Staubli VAL3: tx2.pjx

--- tx2.pjx ---
Parameters version=s8.10.5Cs9_BS2172 stackSize=20000 millimeterUnit=true
Program file=getPath.pgx
Program file=initArmInfo.pgx
Program file=initDataBase.pgx
Program file=initWidget.pgx
Program file=mainCycle.pgx
Program file=moveCalPos.pgx
Program file=moveRecPos.pgx
Program file=refreshBtn0_CaliTcp.pgx
Program file=refreshBtn1_AdjXY.pgx
Program file=refreshBtn2_AdjZ.pgx
Program file=refreshBtn3_Test.pgx
Program file=saveCall.pgx
Program file=saveTask.pgx
Program file=start.pgx
Program file=stop.pgx
Data file=tx2.dtx
Library alias=algorithm path=Disk://SmartTCP_CS9/Algorithm6/Algorithm6.pjx
Library alias=db path=Disk://SmartTCP_CS9/DataBase6/DataBase6.pjx

--- tx2.dtx ---


--- start.pgx ---
public program start()
begin
  call initArmInfo()
  call initWidget()
  call initDataBase()
  call mainCycle()
end

--- getPath.pgx ---
program getPath(string x_sHmiName, string& x_sHmiPath)
begin
  x_sHmiPath=libPath()+"/interface/"+x_sHmiName
end

--- initArmInfo.pgx ---
program initArmInfo()
  local string l_sLanguage
  local string l_sMounting
begin
  //*******************************************************
  db:utLbl_Axis_Data.Common.sText="6axis"
  //*******************************************************
  //Get mounting property
  //*******************************************************
  l_sMounting=getVersion("Arm Mounting")
  switch l_sMounting
    case "floor"
      db:sMounting="Floor"
      db:utCbx_Mounting_Data.Common.sValue="Floor"
    break
    case "ceiling"
      db:sMounting="Ceiling"
      db:utCbx_Mounting_Data.Common.sValue="Ceiling"
    break
    default
      db:sMounting="Null"
      db:utCbx_Mounting_Data.Common.sValue=""
    break
  endSwitch
  //*******************************************************
  //Get system language
  //*******************************************************
  l_sLanguage=getLanguage()
  switch l_sLanguage
    case "chinese"
      db:sLanguage="chinese"
      db:utCbx_Language_Data.Common.sValue="Chinese"
    break
    case "english"
      db:sLanguage="english"
      db:utCbx_Language_Data.Common.sValue="English"
    break
    default
      db:sLanguage="english"
      db:utCbx_Language_Data.Common.sValue="English"
    break
  endSwitch
  //
  //*******************************************************
  //Initialize the flange as the current tool
  //*******************************************************
  call db:updateTool(0,false)
end

--- initDataBase.pgx ---
program initDataBase()
begin
  db:nStep0=10
  db:nStep1=10
  db:nStep2=10
  db:nStep3=10
  //
  db:tFlange.trsf={0,0,0,0,0,0}
  db:trOffset={0,0,10,0,0,0}
  //
  db:mSpeed_C_blend.tvel=250
  db:mSpeed_C_blend.blend=Cartesian
  db:mSpeed_C_blend.leave=0
  db:mSpeed_C_blend.reach=0
  //
  db:mSpeed_J_blend.tvel=250
  db:mSpeed_J_blend.blend=joint
  db:mSpeed_J_blend.leave=5
  db:mSpeed_J_blend.reach=5
  //
  db:mSlow.tvel=30
  db:mSlow.blend=Cartesian
  db:mSlow.leave=0
  db:mSlow.reach=0
  //
  db:cConfigSame={ssame,esame,wsame}
  //
  //pTeach1.trsf={0,0,0,0,0,0}
  db:pTeach1.config={ssame,esame,wsame}
  //pTeach2.trsf={0,0,0,0,0,0}
  db:pTeach2.config={ssame,esame,wsame}
  //pTeach3.trsf={0,0,0,0,0,0}
  db:pTeach3.config={ssame,esame,wsame}
  //pTeach4.trsf={0,0,0,0,0,0}
  db:pTeach4.config={ssame,esame,wsame}
  //pTeach5.trsf={0,0,0,0,0,0}
  db:pTeach5.config={ssame,esame,wsame}
  //pTeach6.trsf={0,0,0,0,0,0}
  db:pTeach6.config={ssame,esame,wsame}
  //pTeach6.trsf={0,0,0,0,0,0}
  db:pTeach7.config={ssame,esame,wsame}
  //
  //pAdjustXY_2_1.trsf={0,0,0,0,0,0}
  db:pAdjustXY_2_1.config={ssame,esame,wsame}
  //pAdjustXY_2_2.trsf={0,0,0,0,0,0}
  db:pAdjustXY_2_2.config={ssame,esame,wsame}
  //pAdjustXY_3_1.trsf={0,0,0,0,0,0}
  db:pAdjustXY_3_1.config={ssame,esame,wsame}
  //pAdjustXY_3_2.trsf={0,0,0,0,0,0}
  db:pAdjustXY_3_2.config={ssame,esame,wsame}
  //pAdjustXY_3_3.trsf={0,0,0,0,0,0}
  db:pAdjustXY_3_3.config={ssame,esame,wsame}
  //pAdjustZ_2_1.trsf={0,0,0,0,0,0}
  db:pAdjustZ_2_1.config={ssame,esame,wsame}
  //pAdjustZ_2_2.trsf={0,0,0,0,0,0}
  db:pAdjustZ_2_2.config={ssame,esame,wsame}
  //
  db:bTeach1=false
  db:bTeach2=false
  db:bTeach3=false
  db:bTeach4=false
  db:bTeach5=false
  db:bTeach6=false
  db:bTeach7=false
  //
  db:bAdjustXY_2_1=false
  db:bAdjustXY_2_2=false
  db:bAdjustXY_3_1=false
  db:bAdjustXY_3_2=false
  db:bAdjustXY_3_3=false
  db:bAdjustZ_2_1=false
  db:bAdjustZ_2_2=false
  //
  db:sLanguageM=""
  db:sCbxLanguage=""
  db:sCbxMounting=""
end

--- initWidget.pgx ---
program initWidget()
  local num l_nI
  local string l_sID
  local string l_sPage
begin
  //*************************************************************************************************
  //Initialize the widgets of the <Page_Main>：
  //*************************************************************************************************
  call getPath("Page_Main",l_sPage)
  //Container
  call db:initContainer(db:utCtn_Function,l_sPage,"ctn_Function",true)
  db:utCtn_Function.Common.sSource="Page_Container_Main.html"
  db:utCtn_Function.Appearance.bVisibility=true
  call db:initContainer(db:utCtn_Message,l_sPage,"ctn_Message",false)
  db:utCtn_Message.Common.sSource="Page_Container_Alert.html"
  db:utCtn_Message.Appearance.bVisibility=false
  //
  //Button
  call db:initButton(db:utBtn_Bottom[0],l_sPage,"bottom_btn0","")
  call db:initButton(db:utBtn_Bottom[1],l_sPage,"bottom_btn1","")
  call db:initButton(db:utBtn_Bottom[2],l_sPage,"bottom_btn2","")
  call db:initButton(db:utBtn_Bottom[3],l_sPage,"bottom_btn3","")
  call db:initButton(db:utBtn_Bottom[4],l_sPage,"bottom_btn4","")
  call db:initButton(db:utBtn_Bottom[5],l_sPage,"bottom_btn5","")
  call db:initButton(db:utBtn_Bottom[6],l_sPage,"bottom_btn6","")
  call db:initButton(db:utBtn_Bottom[7],l_sPage,"bottom_btn7","")
  call db:updateBtn(83,"Null,Null,Null,Null,Null,Null,Null,Quit")
  //
  //Combo
  call db:initCombo(db:utCbx_Language_Data,l_sPage,"cbx_Language_D")
  call db:initCombo(db:utCbx_Mounting_Data,l_sPage,"cbx_Mounting_D")
  //
  //Label
  call db:initLabel(db:utLbl_Title,l_sPage,"lbl_Title","Stäubli Tool Calibration - SmartTCP")
  db:utLbl_Title.Appearance.sBackgroundColour="rgba(0,0,255,0.251)"
  call db:initLabel(db:utLbl_Language,l_sPage,"lbl_Language","Language：")
  //
  call db:initLabel(db:utLbl_Axis,l_sPage,"lbl_Axis","ArmType：")
  call db:initLabel(db:utLbl_Axis_Data,l_sPage,"lbl_Axis_Data","6Axis")
  call db:initLabel(db:utLbl_Mounting,l_sPage,"lbl_Mounting","Mounting：")
  call db:initLabel(db:utLbl_Tool,l_sPage,"lbl_Tool","Tool：")
  call db:initLabel(db:utLbl_Tool_Data,l_sPage,"lbl_Tool_Data","tFlange")
  call db:initLabel(db:utLbl_CurrentPos_Name[0],l_sPage,"lbl_CurrentPos_Name0","X")
  call db:initLabel(db:utLbl_CurrentPos_Name[1],l_sPage,"lbl_CurrentPos_Name1","Y")
  call db:initLabel(db:utLbl_CurrentPos_Name[2],l_sPage,"lbl_CurrentPos_Name2","Z")
  call db:initLabel(db:utLbl_CurrentPos_Name[3],l_sPage,"lbl_CurrentPos_Name3","RX")
  call db:initLabel(db:utLbl_CurrentPos_Name[4],l_sPage,"lbl_CurrentPos_Name4","RY")
  call db:initLabel(db:utLbl_CurrentPos_Name[5],l_sPage,"lbl_CurrentPos_Name5","RZ")
  //
  for l_nI= 0 to 5
    l_sID="lbl_CurrentPos_Data"+toString("0,0",l_nI)
    call db:initLabel(db:utLbl_CurrentPos_Data[l_nI],l_sPage,l_sID,"Null")
  endFor
  //
  call db:initLabel(db:utLbl_Info0,l_sPage,"lbl_info0","Null")
  call db:initLabel(db:utLbl_Info1,l_sPage,"lbl_info1","Null")
  call db:initLabel(db:utLbl_Info2,l_sPage,"lbl_info2","Null")
  call db:initLabel(db:utLbl_Info3,l_sPage,"lbl_info3","Null")
  call db:initLabel(db:utLbl_Info4,l_sPage,"lbl_info4","Null")
  call db:updateInfo(100,db:utLbl_Info2.Data.nVal,db:utLbl_Info2.Common.sText,"0","TCP calibration application for TX2/TS2 robot")
  //
  //Image
  call db:initImage(db:utImg_JogMode[0],l_sPage,"img_None")
  call db:initImage(db:utImg_JogMode[1],l_sPage,"img_Joint")
  call db:initImage(db:utImg_JogMode[2],l_sPage,"img_Frame")
  call db:initImage(db:utImg_JogMode[3],l_sPage,"img_Tool")
  db:utImg_JogMode[0].Common.sSourceImage="images/none.svg"
  db:utImg_JogMode[1].Common.sSourceImage="images/joint.svg"
  db:utImg_JogMode[2].Common.sSourceImage="images/frame.svg"
  db:utImg_JogMode[3].Common.sSourceImage="images/tool.svg"
  //
  call db:initImage(db:utImg_Info,l_sPage,"img_info")
  db:utImg_Info.Common.sSourceImage="images/info.png"
  //
  call db:initImage(db:utImg_PosSwitch,l_sPage,"img_PosSwitch")
  db:utImg_PosSwitch.Common.sSourceImage="images/switch.png"
  //*************************************************************************************************
  //
  //
  //*************************************************************************************************
  //Initialize the widgets of the <Page_Container_Main>：
  //*************************************************************************************************
  call getPath("Page_Container_Main",l_sPage)
  //Label
  call db:initLabel(db:utLbl_CheckBox_a[0],l_sPage,"lbl_CheckBox_a0","3Points")
  call db:initLabel(db:utLbl_CheckBox_a[1],l_sPage,"lbl_CheckBox_a1","4Points")
  call db:initLabel(db:utLbl_CheckBox_a[2],l_sPage,"lbl_CheckBox_a2","7Points")
  call db:initLabel(db:utLbl_CheckBox_b[0],l_sPage,"lbl_CheckBox_b0","2Points180°")
  call db:initLabel(db:utLbl_CheckBox_b[1],l_sPage,"lbl_CheckBox_b1","3Points120°")
  //
  //CheckBox_a
  call db:initCheckBox(db:utImg_CheckBox_a[0],l_sPage,"img_CheckBox_a0","CheckOff")
  call db:initCheckBox(db:utImg_CheckBox_a[1],l_sPage,"img_CheckBox_a1","CheckOn")
  call db:initCheckBox(db:utImg_CheckBox_a[2],l_sPage,"img_CheckBox_a2","CheckOff")
  //
  //CheckBox_b
  call db:initCheckBox(db:utImg_CheckBox_b[0],l_sPage,"img_CheckBox_b0","CheckOn")
  call db:initCheckBox(db:utImg_CheckBox_b[1],l_sPage,"img_CheckBox_b1","CheckOff")
  //
  //Button
  call db:initButton(db:utBtn_Step[0],l_sPage,"step_btn0","Calibration tool")
  call db:initButton(db:utBtn_Step[1],l_sPage,"step_btn1","Correction tool XY")
  call db:initButton(db:utBtn_Step[2],l_sPage,"step_btn2","Correction tool Z")
  call db:initButton(db:utBtn_Step[3],l_sPage,"step_btn3","Verification tool")
  //*************************************************************************************************
  //
  //
  //*************************************************************************************************
  //Initialize the widgets of the <Page_Container_Alert>：
  //*************************************************************************************************
  call getPath("Page_Container_Alert",l_sPage)
  //Text
  call db:initText(db:utTxt_popUpMsg,l_sPage,"txt_popUpMsg","String")
  db:utTxt_popUpMsg.Appearance.sBackgroundColour="#7C95FF"
  //
  //Button
  call db:initButton(db:utBtn_OK,l_sPage,"btn_OK","OK")
  //*************************************************************************************************
  //
  //
  //*************************************************************************************************
  //Initialize the widgets of the <Page_Container_Confirm>：
  //*************************************************************************************************
   call getPath("Page_Container_Confirm",l_sPage)
  //Text
  call db:initText(db:utTxt_popUpMsg,l_sPage,"txt_popUpMsg","String")
  //
  //Button
  call db:initButton(db:utBtn_Yes,l_sPage,"btn_Yes","Yes")
  call db:initButton(db:utBtn_No,l_sPage,"btn_No","No")
  //*************************************************************************************************
  //
  //
  //*************************************************************************************************
  //Initialize interface language
  //*************************************************************************************************
  call db:refreshLanguage()
  call db:updateCurrentPos()
  userPage("Page_Main")
  //*************************************************************************************************
  //
  //
  //*************************************************************************************************
  //Initialize the widgets of the <Page_Container_Teach>：
  //*************************************************************************************************
 call getPath("Page_Container_Teach",l_sPage)
  //Label
  for l_nI=0 to 5
    l_sID="utLbl_PosValue_Data"+toString("0.0",l_nI)
    call db:initLabel(db:utLbl_PosValue_Data[l_nI],l_sPage,l_sID,"Null")
  endFor
  call db:initLabel(db:utLbl_Point,l_sPage,"lbl_Point","Point：P1")
  call db:initLabel(db:utLbl_Step,l_sPage,"lbl_Step","Step：1/3")
  //Image
  call db:initImage(db:utImg_Example,l_sPage,"img_example")
  //*************************************************************************************************
  //
  //
  //*************************************************************************************************
  //Initialize the widgets of the <Page_Container_Test>：
  //*************************************************************************************************
  call getPath("Page_Container_Test",l_sPage)
  //Label
  call db:initLabel(db:utLbl_SwitchTool,l_sPage,"lbl_SwitchTool","Tool Switch：")
  call db:initLabel(db:utLbl_Offset,l_sPage,"lbl_Offset","Tool Offset：")
  for l_nI=0 to 5
    l_sID="utLbl_ToolValue_Data"+toString("0.0",l_nI)
    call db:initLabel(db:utLbl_ToolValue_Data[l_nI],l_sPage,l_sID,"Null")
  endFor
  //
  //Text
  for l_nI=0 to 5
    l_sID="utTxt_OffsetValue_Data"+toString("0.0",l_nI)
    call db:initText(db:utTxt_OffsetValue_Data[l_nI],l_sPage,l_sID,"Num")
    db:utTxt_OffsetValue_Data[l_nI].Appearance.sBackgroundColour="#EEFF00"
  endFor
  //
  //Image
  call db:initImage(db:utImg_Previous,l_sPage,"img_Previous")
  db:utImg_Previous.Common.sSourceImage="images/navigate-previous.svg"
  call db:initImage(db:utImg_Next,l_sPage,"img_Next")
  db:utImg_Next.Common.sSourceImage="images/navigate-next.svg"
  //
  //CheckBox
  call db:initCheckBox(db:utImg_Switch,l_sPage,"img_Switch","SwitchOff")
  //*************************************************************************************************
end

--- mainCycle.pgx ---
public program mainCycle()
  local bool l_bOut
  local string l_sStr
  local num l_nVal
  local bool l_bConfirm
begin
  l_bOut=false
  do
    //*************************************************************************************************
    //Refresh the widgets of the <Page_Container_Main>：
    //*************************************************************************************************
    call db:refreshLanguage()
    call db:refreshCheckBox(db:utImg_CheckBox_a)
    call db:refreshCheckBox(db:utImg_CheckBox_b)
    call db:refreshJogMode()
    call db:refreshInfo()
    call db:refreshQuit(l_bOut)
    //
    call refreshBtn0_CaliTcp()
    //
    call refreshBtn1_AdjXY()
    //
    call refreshBtn2_AdjZ()
    //
    call refreshBtn3_Test()

  until l_bOut
end

--- moveCalPos.pgx ---
program moveCalPos(string x_sTarget)
  local bool l_bTaskStatusErr
begin
  if taskStatus("m")!=-1
    taskKill("m")
  endIf
  if taskStatus("m")==-1
    taskCreate "m",100, db:ListMove(x_sTarget)
  endIf
  l_bTaskStatusErr=watch(taskStatus("m")==150 or taskStatus("m")>1,0.3)
  if l_bTaskStatusErr==true
    taskKill("m")
    call db:hmiAlert("CantMove1","warning")
  endIf
end

--- moveRecPos.pgx ---
program moveRecPos(string x_sTarget)
  local bool l_bTaskStatusErr
begin
  if taskStatus("m")!=-1
    taskKill("m")
  endIf
  if taskStatus("m")==-1
    taskCreate "m",100, db:ListMove(x_sTarget)
  endIf
  l_bTaskStatusErr=watch(taskStatus("m")==150 or taskStatus("m")>1,0.3)
  if l_bTaskStatusErr==true
    taskKill("m")
    call db:hmiAlert("CantMove2","warning")
  endIf
end

--- refreshBtn0_CaliTcp.pgx ---
public program refreshBtn0_CaliTcp()
begin
  if db:utBtn_Step[0].Events.bClick==true
    db:utCtn_Function.Common.sSource="Page_Container_Teach.html"
    //**********************************************************************************************************************************
    //3点法标定TCP
    if db:utImg_CheckBox_a[0].Data.bStatus==true
      switch db:nStep0
        case 10
          call db:updateStr(31,db:utLbl_Point.Common.sText,"Point：P1")
          call db:updateStr(43,db:utLbl_Step.Common.sText,"Step：1/3")
          //
          db:utImg_Example.Common.sSourceImage="images/6AxisTeach_1.png"

          //
          call db:updateTeachPos(db:pTeach1,db:bTeach1)
          //
          call db:updateBtn(80,"Align,Here,Move,Null,Null,Null,Prev.,Next")
          //
          call db:updateInfo(101,db:utLbl_Info0.Data.nVal,db:utLbl_Info0.Common.sText,"0","Operation reminder：")
          call db:updateInfo(102,db:utLbl_Info1.Data.nVal,db:utLbl_Info1.Common.sText,"1","Touch to reference pointer in vertical attitude")
          call db:updateInfo(105,db:utLbl_Info2.Data.nVal,db:utLbl_Info2.Common.sText,"2","Press Here button to save the position")
          call db:updateInfo(125,db:utLbl_Info3.Data.nVal,db:utLbl_Info3.Common.sText,"3","Alignment can be used when the tool and flange are 90°")
          call db:updateInfo(99,db:utLbl_Info4.Data.nVal,db:utLbl_Info4.Common.sText,"4","")
          //
          call db:updateTool(0,false)
          db:nStep0=11
        break
        //
        case 11
          if db:utBtn_Bottom[0].Events.bClick==true
            db:utBtn_Bottom[0].Events.bClick=false
            //Press F1
            call moveCalPos("Align")
          endIf

          if db:utBtn_Bottom[1].Events.bClick==true
            db:utBtn_Bottom[1].Events.bClick=false
            //Press F2
            db:bTeach1=true
            db:pTeach1=here(flange,world)
            db:jTeach1=herej()
            call db:updateTeachPos(db:pTeach1,db:bTeach1)
            call db:hmiAlert("First","info")
            call saveCall()
          endIf
          if db:utBtn_Bottom[2].Events.bClick==true
            db:utBtn_Bottom[2].Events.bClick=false
            //Press F3
            call moveRecPos("pTeach1")
          endIf
          if db:utBtn_Bottom[6].Events.bClick==true
            db:utBtn_Bottom[6].Events.bClick=false
            //Press F7
            resetMotion()
            db:utCtn_Message.Appearance.bVisibility=false
            db:nStep0=99
          endIf
          if db:utBtn_Bottom[7].Events.bClick==true
            db:utBtn_Bottom[7].Events.bClick=false
            //Press F8
            resetMotion()
            db:utCtn_Message.Appearance.bVisibility=false
            db:nStep0=20
          endIf
        break
        //
        case 20
          call db:updateStr(32,db:utLbl_Point.Common.sText,"Point：P2")
          call db:updateStr(44,db:utLbl_Step.Common.sText,"Step：2/3")
          //
          db:utImg_Example.Common.sSourceImage="images/6AxisTeach_2.png"

          //
          call db:updateTeachPos(db:pTeach2,db:bTeach2)
          //
          call db:updateBtn(81,"Null,Here,Move,Null,Null,Null,Prev.,Next")
          //
          call db:updateInfo(101,db:utLbl_Info0.Data.nVal,db:utLbl_Info0.Common.sText,"0","Operation reminder：")
          call db:updateInfo(103,db:utLbl_Info1.Data.nVal,db:utLbl_Info1.Common.sText,"1","Touch to reference pointer in any attitude")
          call db:updateInfo(105,db:utLbl_Info2.Data.nVal,db:utLbl_Info2.Common.sText,"2","Press Here button to save the position")
          call db:updateInfo(99,db:utLbl_Info3.Data.nVal,db:utLbl_Info3.Common.sText,"3","")
          call db:updateInfo(99,db:utLbl_Info4.Data.nVal,db:utLbl_Info4.Common.sText,"4","")
          db:nStep0=21
        break
        //
        case 21
          if db:utBtn_Bottom[1].Events.bClick==true
            db:utBtn_Bottom[1].Events.bClick=false
            //Press F2
            db:bTeach2=true
            db:pTeach2=here(flange,world)
            db:jTeach2=herej()
            call db:updateTeachPos(db:pTeach2,db:bTeach2)
            call db:hmiAlert("Second","info")
            call saveCall()
          endIf
          if db:utBtn_Bottom[2].Events.bClick==true
            db:utBtn_Bottom[2].Events.bClick=false
            //Press F3
            call moveRecPos("pTeach2")
          endIf
          if db:utBtn_Bottom[6].Events.bClick==true
            db:utBtn_Bottom[6].Events.bClick=false
            //Press F7
            resetMotion()
            db:utCtn_Message.Appearance.bVisibility=false
            db:nStep0=10
          endIf
          if db:utBtn_Bottom[7].Events.bClick==true
            db:utBtn_Bottom[7].Events.bClick=false
            //Press F8
            resetMotion()
            db:utCtn_Message.Appearance.bVisibility=false
            db:nStep0=30
          endIf
        break
        //
        case 30
          call db:updateStr(33,db:utLbl_Point.Common.sText,"Point：P3")
          call db:updateStr(45,db:utLbl_Step.Common.sText,"Step：3/3")
          //
          db:utImg_Example.Common.sSourceImage="images/6AxisTeach_3.png"

          //
          call db:updateTeachPos(db:pTeach3,db:bTeach3)
          //
          call db:updateBtn(82,"Null,Here,Move,Null,Null,Calc.,Prev.,Done")
          //
          call db:updateInfo(101,db:utLbl_Info0.Data.nVal,db:utLbl_Info0.Common.sText,"0","Operation reminder：")
          call db:updateInfo(103,db:utLbl_Info1.Data.nVal,db:utLbl_Info1.Common.sText,"1","Touch to reference pointer in any attitude")
          call db:updateInfo(105,db:utLbl_Info2.Data.nVal,db:utLbl_Info2.Common.sText,"2","Press Here button to save the position")
          call db:updateInfo(104,db:utLbl_Info3.Data.nVal,db:utLbl_Info3.Common.sText,"3","Press Calc. button to get the TCP value")
          call db:updateInfo(99,db:utLbl_Info4.Data.nVal,db:utLbl_Info4.Common.sText,"4","")
          db:nStep0=31
        break
        //
        case 31
          if db:utBtn_Bottom[1].Events.bClick==true
            db:utBtn_Bottom[1].Events.bClick=false
            //Press F2
            db:bTeach3=true
            db:pTeach3=here(flange,world)
            db:jTeach3=herej()
            call db:updateTeachPos(db:pTeach3,db:bTeach3)
            call db:hmiAlert("Third","info")
            call saveCall()
          endIf
          if db:utBtn_Bottom[2].Events.bClick==true
            db:utBtn_Bottom[2].Events.bClick=false
            //Press F3
            call moveRecPos("pTeach3")
          endIf
          if db:utBtn_Bottom[5].Events.bClick==true
            db:utBtn_Bottom[5].Events.bClick=false
            //Press F6
            call algorithm:CalToolPos3(db:tTool1)
          endIf
          if db:utBtn_Bottom[6].Events.bClick==true
            db:utBtn_Bottom[6].Events.bClick=false
            //Press F7
            resetMotion()
            db:utCtn_Message.Appearance.bVisibility=false
            db:nStep0=20
          endIf
          if db:utBtn_Bottom[7].Events.bClick==true
            db:utBtn_Bottom[7].Events.bClick=false
            //Press F8
            resetMotion()
            db:utCtn_Message.Appearance.bVisibility=false
            db:nStep0=99
          endIf
        break
        //
        case 99
          db:utCtn_Function.Common.sSource="Page_Container_Main.html"
          //
          call db:updateBtn(83,"Null,Null,Null,Null,Null,Null,Null,Quit")
          //
          call db:updateInfo(99,db:utLbl_Info0.Data.nVal,db:utLbl_Info0.Common.sText,"0","")
          call db:updateInfo(99,db:utLbl_Info1.Data.nVal,db:utLbl_Info1.Common.sText,"1","")
          call db:updateInfo(100,db:utLbl_Info2.Data.nVal,db:utLbl_Info2.Common.sText,"0","TCP calibration application for TX2/TS2 robot")
          call db:updateInfo(99,db:utLbl_Info3.Data.nVal,db:utLbl_Info3.Common.sText,"3","")
          call db:updateInfo(99,db:utLbl_Info4.Data.nVal,db:utLbl_Info4.Common.sText,"4","")
          db:utBtn_Step[0].Events.bClick=false
          db:nStep0=10
        break
        //
      endSwitch
    endIf
    //**********************************************************************************************************************************
    //
    //**********************************************************************************************************************************
    //4点法标定TCP
    if db:utImg_CheckBox_a[1].Data.bStatus==true
      switch db:nStep0
        case 10

          call db:updateStr(31,db:utLbl_Point.Common.sText,"Point：P1")
          call db:updateStr(46,db:utLbl_Step.Common.sText,"Step：1/4")
          //
          db:utImg_Example.Common.sSourceImage="images/6AxisTeach_1.png"

          //
          call db:updateTeachPos(db:pTeach1,db:bTeach1)
          //
          call db:updateBtn(80,"Align,Here,Move,Null,Null,Null,Prev.,Next")
          //
          call db:updateInfo(101,db:utLbl_Info0.Data.nVal,db:utLbl_Info0.Common.sText,"0","Operation reminder：")
          call db:updateInfo(102,db:utLbl_Info1.Data.nVal,db:utLbl_Info1.Common.sText,"1","Touch to reference pointer in vertical attitude")
          call db:updateInfo(105,db:utLbl_Info2.Data.nVal,db:utLbl_Info2.Common.sText,"2","Press Here button to save the position")
          call db:updateInfo(125,db:utLbl_Info3.Data.nVal,db:utLbl_Info3.Common.sText,"3","Alignment can be used when the tool and flange are 90°")
          call db:updateInfo(99,db:utLbl_Info4.Data.nVal,db:utLbl_Info4.Common.sText,"4","")
          //
          call db:updateTool(0,false)
          db:nStep0=11
        break
        //
        case 11
          if db:utBtn_Bottom[0].Events.bClick==true
            db:utBtn_Bottom[0].Events.bClick=false
            //Press F1
            call moveCalPos("Align")
          endIf
          if db:utBtn_Bottom[1].Events.bClick==true
            db:utBtn_Bottom[1].Events.bClick=false
            //Press F2
            db:bTeach1=true
            db:pTeach1=here(flange,world)
            db:jTeach1=herej()
            call db:updateTeachPos(db:pTeach1,db:bTeach1)
            call db:hmiAlert("First","info")
            call saveCall()
          endIf
          if db:utBtn_Bottom[2].Events.bClick==true
            db:utBtn_Bottom[2].Events.bClick=false
            //Press F3
            call moveRecPos("pTeach1")
          endIf
          if db:utBtn_Bottom[6].Events.bClick==true
            db:utBtn_Bottom[6].Events.bClick=false
            //Press F7
            resetMotion()
            db:utCtn_Message.Appearance.bVisibility=false
            db:nStep0=99
          endIf
          if db:utBtn_Bottom[7].Events.bClick==true
            db:utBtn_Bottom[7].Events.bClick=false
            //Press F8
            resetMotion()
            db:utCtn_Message.Appearance.bVisibility=false
            db:nStep0=20
          endIf
        break
        //
        case 20
          call db:updateStr(32,db:utLbl_Point.Common.sText,"Point：P2")
          call db:updateStr(47,db:utLbl_Step.Common.sText,"Step：2/4")
          //
          db:utImg_Example.Common.sSourceImage="images/6AxisTeach_2.png"

          //
          call db:updateTeachPos(db:pTeach2,db:bTeach2)
          //
          call db:updateBtn(81,"Null,Here,Move,Null,Null,Null,Prev.,Next")
          //
          call db:updateInfo(101,db:utLbl_Info0.Data.nVal,db:utLbl_Info0.Common.sText,"0","Operation reminder：")
          call db:updateInfo(103,db:utLbl_Info1.Data.nVal,db:utLbl_Info1.Common.sText,"1","Touch to reference pointer in any attitude")
          call db:updateInfo(105,db:utLbl_Info2.Data.nVal,db:utLbl_Info2.Common.sText,"2","Press Here button to save the position")
          call db:updateInfo(99,db:utLbl_Info3.Data.nVal,db:utLbl_Info3.Common.sText,"3","")
          call db:updateInfo(99,db:utLbl_Info4.Data.nVal,db:utLbl_Info4.Common.sText,"4","")
          db:nStep0=21
        break
        //
        case 21
          if db:utBtn_Bottom[1].Events.bClick==true
            db:utBtn_Bottom[1].Events.bClick=false
            //Press F2
            db:bTeach2=true
            db:pTeach2=here(flange,world)
            db:jTeach2=herej()
            call db:updateTeachPos(db:pTeach2,db:bTeach2)
            call db:hmiAlert("Second","info")
            call saveCall()
          endIf
          if db:utBtn_Bottom[2].Events.bClick==true
            db:utBtn_Bottom[2].Events.bClick=false
            //Press F3
            call moveRecPos("pTeach2")
          endIf
          if db:utBtn_Bottom[6].Events.bClick==true
            db:utBtn_Bottom[6].Events.bClick=false
            //Press F7
            resetMotion()
            db:utCtn_Message.Appearance.bVisibility=false
            db:nStep0=10
          endIf
          if db:utBtn_Bottom[7].Events.bClick==true
            db:utBtn_Bottom[7].Events.bClick=false
            //Press F8
            resetMotion()
            db:utCtn_Message.Appearance.bVisibility=false
            db:nStep0=30
          endIf
        break
        //
        case 30
          call db:updateStr(33,db:utLbl_Point.Common.sText,"Point：P3")
          call db:updateStr(48,db:utLbl_Step.Common.sText,"Step：3/4")
          //
          db:utImg_Example.Common.sSourceImage="images/6AxisTeach_3.png"

          //
          call db:updateTeachPos(db:pTeach3,db:bTeach3)
          //
          call db:updateBtn(81,"Null,Here,Move,Null,Null,Null,Prev.,Next")
          //
          call db:updateInfo(101,db:utLbl_Info0.Data.nVal,db:utLbl_Info0.Common.sText,"0","Operation reminder：")
          call db:updateInfo(103,db:utLbl_Info1.Data.nVal,db:utLbl_Info1.Common.sText,"1","Touch to reference pointer in any attitude")
          call db:updateInfo(105,db:utLbl_Info2.Data.nVal,db:utLbl_Info2.Common.sText,"2","Press Here button to save the position")
          call db:updateInfo(99,db:utLbl_Info3.Data.nVal,db:utLbl_Info3.Common.sText,"3","")
          call db:updateInfo(99,db:utLbl_Info4.Data.nVal,db:utLbl_Info4.Common.sText,"4","")
          db:nStep0=31
        break
        //
        case 31
          if db:utBtn_Bottom[1].Events.bClick==true
            db:utBtn_Bottom[1].Events.bClick=false
            //Press F2
            db:bTeach3=true
            db:pTeach3=here(flange,world)
            db:jTeach3=herej()
            call db:updateTeachPos(db:pTeach3,db:bTeach3)
            call db:hmiAlert("Third","info")
            call saveCall()
          endIf
          if db:utBtn_Bottom[2].Events.bClick==true
            db:utBtn_Bottom[2].Events.bClick=false
            //Press F3
            call moveRecPos("pTeach3")
          endIf
          if db:utBtn_Bottom[6].Events.bClick==true
            db:utBtn_Bottom[6].Events.bClick=false
            //Press F7
            resetMotion()
            db:utCtn_Message.Appearance.bVisibility=false
            db:nStep0=20
          endIf
          if db:utBtn_Bottom[7].Events.bClick==true
            db:utBtn_Bottom[7].Events.bClick=false
            //Press F8
            resetMotion()
            db:utCtn_Message.Appearance.bVisibility=false
            db:nStep0=40
          endIf
        break
        //
        case 40
          call db:updateStr(34,db:utLbl_Point.Common.sText,"Point：P4")
          call db:updateStr(49,db:utLbl_Step.Common.sText,"Step：4/4")
          //
          db:utImg_Example.Common.sSourceImage="images/6AxisTeach_4.png"

          //
          call db:updateTeachPos(db:pTeach4,db:bTeach4)
          //
          call db:updateBtn(82,"Null,Here,Move,Null,Null,Calc.,Prev.,Done")
          //
          call db:updateInfo(101,db:utLbl_Info0.Data.nVal,db:utLbl_Info0.Common.sText,"0","Operation reminder：")
          call db:updateInfo(103,db:utLbl_Info1.Data.nVal,db:utLbl_Info1.Common.sText,"1","Touch to reference pointer in any attitude")
          call db:updateInfo(105,db:utLbl_Info2.Data.nVal,db:utLbl_Info2.Common.sText,"2","Press Here button to save the position")
          call db:updateInfo(104,db:utLbl_Info3.Data.nVal,db:utLbl_Info3.Common.sText,"3","Press Calc. button to get the TCP value")
          call db:updateInfo(99,db:utLbl_Info4.Data.nVal,db:utLbl_Info4.Common.sText,"4","")
          db:nStep0=41
        break
        //
        case 41
          if db:utBtn_Bottom[1].Events.bClick==true
            db:utBtn_Bottom[1].Events.bClick=false
            //Press F2
            db:bTeach4=true
            db:pTeach4=here(flange,world)
            db:jTeach4=herej()
            call db:updateTeachPos(db:pTeach4,db:bTeach4)
            call db:hmiAlert("Fourth","info")
            call saveCall()
          endIf
          if db:utBtn_Bottom[2].Events.bClick==true
            db:utBtn_Bottom[2].Events.bClick=false
            //Press F3
            call moveRecPos("pTeach4")
          endIf
          if db:utBtn_Bottom[5].Events.bClick==true
            db:utBtn_Bottom[5].Events.bClick=false
            //Press F6
            call algorithm:CalToolPos4(db:tTool1)
          endIf
          if db:utBtn_Bottom[6].Events.bClick==true
            db:utBtn_Bottom[6].Events.bClick=false
            //Press F7
            resetMotion()
            db:utCtn_Message.Appearance.bVisibility=false
            db:nStep0=30
          endIf
          if db:utBtn_Bottom[7].Events.bClick==true
            db:utBtn_Bottom[7].Events.bClick=false
            //Press F8
            resetMotion()
            db:utCtn_Message.Appearance.bVisibility=false
            db:nStep0=99
          endIf
        break
        //
        case 99
          db:utCtn_Function.Common.sSource="Page_Container_Main.html"
          //
          call db:updateBtn(83,"Null,Null,Null,Null,Null,Null,Null,Quit")
          //
          call db:updateInfo(99,db:utLbl_Info0.Data.nVal,db:utLbl_Info0.Common.sText,"0","")
          call db:updateInfo(99,db:utLbl_Info1.Data.nVal,db:utLbl_Info1.Common.sText,"1","")
          call db:updateInfo(100,db:utLbl_Info2.Data.nVal,db:utLbl_Info2.Common.sText,"0","TCP calibration application for TX2/TS2 robot")
          call db:updateInfo(99,db:utLbl_Info3.Data.nVal,db:utLbl_Info3.Common.sText,"3","")
          call db:updateInfo(99,db:utLbl_Info4.Data.nVal,db:utLbl_Info4.Common.sText,"4","")
          db:utBtn_Step[0].Events.bClick=false
          db:nStep0=10
        break
        //
      endSwitch
    endIf
    //**********************************************************************************************************************************
    //
    //**********************************************************************************************************************************
    //7点法标定TCP
    if db:utImg_CheckBox_a[2].Data.bStatus==true
      switch db:nStep0
        case 10
          call db:updateStr(31,db:utLbl_Point.Common.sText,"Point：P1")
          call db:updateStr(50,db:utLbl_Step.Common.sText,"Step：1/7")
          //
          db:utImg_Example.Common.sSourceImage="images/6AxisTeach_1.png"

          //
          call db:updateTeachPos(db:pTeach1,db:bTeach1)
          //
          call db:updateBtn(80,"Align,Here,Move,Null,Null,Null,Prev.,Next")
          //
          call db:updateInfo(101,db:utLbl_Info0.Data.nVal,db:utLbl_Info0.Common.sText,"0","Operation reminder：")
          call db:updateInfo(102,db:utLbl_Info1.Data.nVal,db:utLbl_Info1.Common.sText,"1","Touch to reference pointer in vertical attitude")
          call db:updateInfo(105,db:utLbl_Info2.Data.nVal,db:utLbl_Info2.Common.sText,"2","Press Here button to save the position")
          call db:updateInfo(125,db:utLbl_Info3.Data.nVal,db:utLbl_Info3.Common.sText,"3","Alignment can be used when the tool and flange are 90°")
          call db:updateInfo(99,db:utLbl_Info4.Data.nVal,db:utLbl_Info4.Common.sText,"4","")
          //
          call db:updateTool(0,false)
          db:nStep0=11
        break
        //
        case 11
          if db:utBtn_Bottom[0].Events.bClick==true
            db:utBtn_Bottom[0].Events.bClick=false
            //Press F1
            call moveCalPos("Align")
          endIf
          if db:utBtn_Bottom[1].Events.bClick==true
            db:utBtn_Bottom[1].Events.bClick=false
            //Press F2
            db:bTeach1=true
            db:pTeach1=here(flange,world)
            db:jTeach1=herej()
            call db:updateTeachPos(db:pTeach1,db:bTeach1)
            call db:hmiAlert("First","info")
            call saveCall()
          endIf
          if db:utBtn_Bottom[2].Events.bClick==true
            db:utBtn_Bottom[2].Events.bClick=false
            //Press F3
            call moveRecPos("pTeach1")
          endIf
          if db:utBtn_Bottom[6].Events.bClick==true
            db:utBtn_Bottom[6].Events.bClick=false
            //Press F7
            resetMotion()
            db:utCtn_Message.Appearance.bVisibility=false
            db:nStep0=99
          endIf
          if db:utBtn_Bottom[7].Events.bClick==true
            db:utBtn_Bottom[7].Events.bClick=false
            //Press F8
            resetMotion()
            db:utCtn_Message.Appearance.bVisibility=false
            db:nStep0=20
          endIf
        break
        //
        case 20
          call db:updateStr(32,db:utLbl_Point.Common.sText,"Point：P2")
          call db:updateStr(51,db:utLbl_Step.Common.sText,"Step：2/7")
          //
          db:utImg_Example.Common.sSourceImage="images/6AxisTeach_2.png"

          //
          call db:updateTeachPos(db:pTeach2,db:bTeach2)
          //
          call db:updateBtn(81,"Null,Here,Move,Null,Null,Null,Prev.,Next")
          //
          call db:updateInfo(101,db:utLbl_Info0.Data.nVal,db:utLbl_Info0.Common.sText,"0","Operation reminder：")
          call db:updateInfo(103,db:utLbl_Info1.Data.nVal,db:utLbl_Info1.Common.sText,"1","Touch to reference pointer in any attitude")
          call db:updateInfo(105,db:utLbl_Info2.Data.nVal,db:utLbl_Info2.Common.sText,"2","Press Here button to save the position")
          call db:updateInfo(99,db:utLbl_Info3.Data.nVal,db:utLbl_Info3.Common.sText,"3","")
          call db:updateInfo(99,db:utLbl_Info4.Data.nVal,db:utLbl_Info4.Common.sText,"4","")
          db:nStep0=21
        break
        //
        case 21
          if db:utBtn_Bottom[1].Events.bClick==true
            db:utBtn_Bottom[1].Events.bClick=false
            //Press F2
            db:bTeach2=true
            db:pTeach2=here(flange,world)
            db:jTeach2=herej()
            call db:updateTeachPos(db:pTeach2,db:bTeach2)
            call db:hmiAlert("Second","info")
            call saveCall()
          endIf
          if db:utBtn_Bottom[2].Events.bClick==true
            db:utBtn_Bottom[2].Events.bClick=false
            //Press F3
            call moveRecPos("pTeach2")
          endIf
          if db:utBtn_Bottom[6].Events.bClick==true
            db:utBtn_Bottom[6].Events.bClick=false
            //Press F7
            resetMotion()
            db:utCtn_Message.Appearance.bVisibility=false
            db:nStep0=10
          endIf
          if db:utBtn_Bottom[7].Events.bClick==true
            db:utBtn_Bottom[7].Events.bClick=false
            //Press F8
            resetMotion()
            db:utCtn_Message.Appearance.bVisibility=false
            db:nStep0=30
          endIf
        break
        //
        case 30
          call db:updateStr(33,db:utLbl_Point.Common.sText,"Point：P3")
          call db:updateStr(52,db:utLbl_Step.Common.sText,"Step：3/7")
          //
          db:utImg_Example.Common.sSourceImage="images/6AxisTeach_3.png"

          //
          call db:updateTeachPos(db:pTeach3,db:bTeach3)
          //
          call db:updateBtn(81,"Null,Here,Move,Null,Null,Null,Prev.,Next")
          //
          call db:updateInfo(101,db:utLbl_Info0.Data.nVal,db:utLbl_Info0.Common.sText,"0","Operation reminder：")
          call db:updateInfo(103,db:utLbl_Info1.Data.nVal,db:utLbl_Info1.Common.sText,"1","Touch to reference pointer in any attitude")
          call db:updateInfo(105,db:utLbl_Info2.Data.nVal,db:utLbl_Info2.Common.sText,"2","Press Here button to save the position")
          call db:updateInfo(99,db:utLbl_Info3.Data.nVal,db:utLbl_Info3.Common.sText,"3","")
          call db:updateInfo(99,db:utLbl_Info4.Data.nVal,db:utLbl_Info4.Common.sText,"4","")
          db:nStep0=31
        break
        //
        case 31
          if db:utBtn_Bottom[1].Events.bClick==true
            db:utBtn_Bottom[1].Events.bClick=false
            //Press F2
            db:bTeach3=true
            db:pTeach3=here(flange,world)
            db:jTeach3=herej()
            call db:updateTeachPos(db:pTeach3,db:bTeach3)
            call db:hmiAlert("Third","info")
            call saveCall()
          endIf
          if db:utBtn_Bottom[2].Events.bClick==true
            db:utBtn_Bottom[2].Events.bClick=false
            //Press F3
            call moveRecPos("pTeach3")
          endIf
          if db:utBtn_Bottom[6].Events.bClick==true
            db:utBtn_Bottom[6].Events.bClick=false
            //Press F7
            resetMotion()
            db:utCtn_Message.Appearance.bVisibility=false
            db:nStep0=20
          endIf
          if db:utBtn_Bottom[7].Events.bClick==true
            db:utBtn_Bottom[7].Events.bClick=false
            //Press F8
            resetMotion()
            db:utCtn_Message.Appearance.bVisibility=false
            db:nStep0=40
          endIf
        break
        //
        case 40
          call db:updateStr(34,db:utLbl_Point.Common.sText,"Point：P4")
          call db:updateStr(53,db:utLbl_Step.Common.sText,"Step：4/7")
          //
          db:utImg_Example.Common.sSourceImage="images/6AxisTeach_4.png"

          //
          call db:updateTeachPos(db:pTeach4,db:bTeach4)
          //
          call db:updateBtn(81,"Null,Here,Move,Null,Null,Null,Prev.,Next")
          //
          call db:updateInfo(101,db:utLbl_Info0.Data.nVal,db:utLbl_Info0.Common.sText,"0","Operation reminder：")
          call db:updateInfo(103,db:utLbl_Info1.Data.nVal,db:utLbl_Info1.Common.sText,"1","Touch to reference pointer in any attitude")
          call db:updateInfo(105,db:utLbl_Info2.Data.nVal,db:utLbl_Info2.Common.sText,"2","Press Here button to save the position")
          call db:updateInfo(99,db:utLbl_Info3.Data.nVal,db:utLbl_Info3.Common.sText,"3","")
          call db:updateInfo(99,db:utLbl_Info4.Data.nVal,db:utLbl_Info4.Common.sText,"4","")
          db:nStep0=41
        break
        //
        case 41
          if db:utBtn_Bottom[1].Events.bClick==true
            db:utBtn_Bottom[1].Events.bClick=false
            //Press F2
            db:bTeach4=true
            db:pTeach4=here(flange,world)
            db:jTeach4=herej()
            call db:updateTeachPos(db:pTeach4,db:bTeach4)
            call db:hmiAlert("Fourth","info")
            call saveCall()
          endIf
          if db:utBtn_Bottom[2].Events.bClick==true
            db:utBtn_Bottom[2].Events.bClick=false
            //Press F3
            call moveRecPos("pTeach4")
          endIf
          if db:utBtn_Bottom[6].Events.bClick==true
            db:utBtn_Bottom[6].Events.bClick=false
            //Press F7
            resetMotion()
            db:utCtn_Message.Appearance.bVisibility=false
            db:nStep0=30
          endIf
          if db:utBtn_Bottom[7].Events.bClick==true
            db:utBtn_Bottom[7].Events.bClick=false
            //Press F8
            call algorithm:CalToolPos4(db:tTool1)
            call db:updateTool(1,false)
            resetMotion()
            db:utCtn_Message.Appearance.bVisibility=false
            db:nStep0=50
          endIf
        break
        //
        case 50
          call db:updateStr(35,db:utLbl_Point.Common.sText,"Point：P5")
          call db:updateStr(54,db:utLbl_Step.Common.sText,"Step：5/7")
          //
          db:utImg_Example.Common.sSourceImage="images/6AxisTeach_5.png"

          //
          call db:updateTeachPos(db:pTeach5,db:bTeach5)
          //
          call db:updateBtn(80,"Align,Here,Move,Null,Null,Null,Prev.,Next")
          //
          call db:updateInfo(101,db:utLbl_Info0.Data.nVal,db:utLbl_Info0.Common.sText,"0","Operation reminder：")
          call db:updateInfo(102,db:utLbl_Info1.Data.nVal,db:utLbl_Info1.Common.sText,"1","Touch to reference pointer in vertical attitude")
          call db:updateInfo(106,db:utLbl_Info2.Data.nVal,db:utLbl_Info2.Common.sText,"2","Press Here button to save the position (Frame Origin)")
          call db:updateInfo(99,db:utLbl_Info3.Data.nVal,db:utLbl_Info3.Common.sText,"3","")
          call db:updateInfo(99,db:utLbl_Info4.Data.nVal,db:utLbl_Info4.Common.sText,"4","")
          db:nStep0=51
        break
        //
        case 51
          if db:utBtn_Bottom[0].Events.bClick==true
            db:utBtn_Bottom[0].Events.bClick=false
            //Press F1
            call moveCalPos("Align")
          endIf
          if db:utBtn_Bottom[1].Events.bClick==true
            db:utBtn_Bottom[1].Events.bClick=false
            //Press F2
            db:bTeach5=true
            db:pTeach5=here(flange,world)
            db:jTeach5=herej()
            call db:updateTeachPos(db:pTeach5,db:bTeach5)
            call db:hmiAlert("Fifth","info")
            call saveCall()
          endIf
          if db:utBtn_Bottom[2].Events.bClick==true
            db:utBtn_Bottom[2].Events.bClick=false
            //Press F3
            call moveRecPos("pTeach5")
          endIf
          if db:utBtn_Bottom[6].Events.bClick==true
            db:utBtn_Bottom[6].Events.bClick=false
            call db:updateTool(0,false)
            resetMotion()
            db:utCtn_Message.Appearance.bVisibility=false
            db:nStep0=40
          endIf
          if db:utBtn_Bottom[7].Events.bClick==true
            db:utBtn_Bottom[7].Events.bClick=false
            resetMotion()
            db:utCtn_Message.Appearance.bVisibility=false
            db:nStep0=60
          endIf
        break
        //
        case 60
          call db:updateStr(36,db:utLbl_Point.Common.sText,"Point：P6")
          call db:updateStr(55,db:utLbl_Step.Common.sText,"Step：6/7")
          //
          db:utImg_Example.Common.sSourceImage="images/6AxisTeach_6.png"

          //
          call db:updateTeachPos(db:pTeach6,db:bTeach6)
          //
          call db:updateBtn(81,"Null,Here,Move,Null,Null,Null,Prev.,Next")
          //
          call db:updateInfo(101,db:utLbl_Info0.Data.nVal,db:utLbl_Info0.Common.sText,"0","Operation reminder：")
          call db:updateInfo(109,db:utLbl_Info1.Data.nVal,db:utLbl_Info1.Common.sText,"1","Keep the current attitude moving in X direction")
          call db:updateInfo(107,db:utLbl_Info2.Data.nVal,db:utLbl_Info2.Common.sText,"2","Press Here button to save the position (Frame Axis OX)")
          call db:updateInfo(99,db:utLbl_Info3.Data.nVal,db:utLbl_Info3.Common.sText,"3","")
          call db:updateInfo(99,db:utLbl_Info4.Data.nVal,db:utLbl_Info4.Common.sText,"4","")
          db:nStep0=61
        break
        //
        case 61
          if db:utBtn_Bottom[1].Events.bClick==true
            db:utBtn_Bottom[1].Events.bClick=false
            //Press F2
            db:bTeach6=true
            db:pTeach6=here(flange,world)
            db:jTeach6=herej()
            call db:updateTeachPos(db:pTeach6,db:bTeach6)
            call db:hmiAlert("Sixth","info")
            call saveCall()
          endIf
          if db:utBtn_Bottom[2].Events.bClick==true
            db:utBtn_Bottom[2].Events.bClick=false
            //Press F3
            call moveRecPos("pTeach6")
          endIf
          if db:utBtn_Bottom[6].Events.bClick==true
            db:utBtn_Bottom[6].Events.bClick=false
            resetMotion()
            db:utCtn_Message.Appearance.bVisibility=false
            db:nStep0=50
          endIf
          if db:utBtn_Bottom[7].Events.bClick==true
            db:utBtn_Bottom[7].Events.bClick=false
            resetMotion()
            db:utCtn_Message.Appearance.bVisibility=false
            db:nStep0=70
          endIf
        break
        //
        case 70
          call db:updateStr(37,db:utLbl_Point.Common.sText,"Point：P7")
          call db:updateStr(56,db:utLbl_Step.Common.sText,"Step：7/7")
          //
          db:utImg_Example.Common.sSourceImage="images/6AxisTeach_7.png"

          //
          call db:updateTeachPos(db:pTeach7,db:bTeach7)
          //
          call db:updateBtn(82,"Null,Here,Move,Null,Null,Calc.,Prev.,Done")
          //
          call db:updateInfo(101,db:utLbl_Info0.Data.nVal,db:utLbl_Info0.Common.sText,"0","Operation reminder：")
          call db:updateInfo(110,db:utLbl_Info1.Data.nVal,db:utLbl_Info1.Common.sText,"1","Keep the current attitude moving in Y direction")
          call db:updateInfo(108,db:utLbl_Info2.Data.nVal,db:utLbl_Info2.Common.sText,"2","Press Here button to save the position (Frame Plane OXY)")
          call db:updateInfo(104,db:utLbl_Info3.Data.nVal,db:utLbl_Info3.Common.sText,"3","Press Calc. button to get the TCP value")
          call db:updateInfo(99,db:utLbl_Info4.Data.nVal,db:utLbl_Info4.Common.sText,"4","")
          db:nStep0=71
        break
        //
        case 71
          if db:utBtn_Bottom[1].Events.bClick==true
            db:utBtn_Bottom[1].Events.bClick=false
            //Press F2
            db:bTeach7=true
            db:pTeach7=here(flange,world)
            db:jTeach7=herej()
            call db:updateTeachPos(db:pTeach7,db:bTeach7)
            call db:hmiAlert("Seventh","info")
            call saveCall()
          endIf
          if db:utBtn_Bottom[2].Events.bClick==true
            db:utBtn_Bottom[2].Events.bClick=false
            //Press F3
            call moveRecPos("pTeach7")
          endIf
          if db:utBtn_Bottom[5].Events.bClick==true
            db:utBtn_Bottom[5].Events.bClick=false
            //Press F6
            call algorithm:CalToolPos7(db:tTool1)
          endIf
          if db:utBtn_Bottom[6].Events.bClick==true
            db:utBtn_Bottom[6].Events.bClick=false
            resetMotion()
            db:utCtn_Message.Appearance.bVisibility=false
            db:nStep0=60
          endIf
          if db:utBtn_Bottom[7].Events.bClick==true
            db:utBtn_Bottom[7].Events.bClick=false
            resetMotion()
            db:utCtn_Message.Appearance.bVisibility=false
            db:nStep0=99
          endIf
        break
        //
        case 99
          db:utCtn_Function.Common.sSource="Page_Container_Main.html"
          //
          call db:updateBtn(83,"Null,Null,Null,Null,Null,Null,Null,Quit")
          //
          call db:updateInfo(99,db:utLbl_Info0.Data.nVal,db:utLbl_Info0.Common.sText,"0","")
          call db:updateInfo(99,db:utLbl_Info1.Data.nVal,db:utLbl_Info1.Common.sText,"1","")
          call db:updateInfo(100,db:utLbl_Info2.Data.nVal,db:utLbl_Info2.Common.sText,"0","TCP calibration application for TX2/TS2 robot")
          call db:updateInfo(99,db:utLbl_Info3.Data.nVal,db:utLbl_Info3.Common.sText,"3","")
          call db:updateInfo(99,db:utLbl_Info4.Data.nVal,db:utLbl_Info4.Common.sText,"4","")
          db:utBtn_Step[0].Events.bClick=false
          db:nStep0=10
        break
        //
      endSwitch
    endIf
    //**********************************************************************************************************************************
  endIf
end

--- refreshBtn1_AdjXY.pgx ---
public program refreshBtn1_AdjXY()
begin
  if db:utBtn_Step[1].Events.bClick==true
    db:utCtn_Function.Common.sSource="Page_Container_Teach.html"
    //**********************************************************************************************************************************
    //2点法修正TCP的XY
    if db:utImg_CheckBox_b[0].Data.bStatus==true
      switch db:nStep1
        case 10
          call db:updateStr(31,db:utLbl_Point.Common.sText,"Point：P1")
          call db:updateStr(41,db:utLbl_Step.Common.sText,"Step：1/2")
          //
          db:utImg_Example.Common.sSourceImage="images/6AxisAdjustXY2_1.png"
          //
          call db:updateTeachPos(db:pAdjustXY_2_1,db:bAdjustXY_2_1)
          //
          call db:updateBtn(84,"Align,Here,Move,Change,Null,Null,Prev.,Next")
          //
          call db:updateInfo(101,db:utLbl_Info0.Data.nVal,db:utLbl_Info0.Common.sText,"0","Operation reminder：")
          call db:updateInfo(113,db:utLbl_Info1.Data.nVal,db:utLbl_Info1.Common.sText,"1","Rotate TCP (RZ) close to one side limit")
          call db:updateInfo(102,db:utLbl_Info2.Data.nVal,db:utLbl_Info2.Common.sText,"2","Touch to reference pointer in vertical attitude")
          call db:updateInfo(111,db:utLbl_Info3.Data.nVal,db:utLbl_Info3.Common.sText,"3","Ensure that the Tool (RZ) reverse can be rotated 180°")
          call db:updateInfo(105,db:utLbl_Info4.Data.nVal,db:utLbl_Info4.Common.sText,"4","Press Here button to save the position")
          //
          call db:updateTool(1,false)
          db:nStep1=11
        break
        //
        case 11
          if db:utBtn_Bottom[0].Events.bClick==true
            db:utBtn_Bottom[0].Events.bClick=false
            //Press F1
            call moveCalPos("Align")
          endIf
          if db:utBtn_Bottom[1].Events.bClick==true
            db:utBtn_Bottom[1].Events.bClick=false
            //Press F2
            db:bAdjustXY_2_1=true
            db:pAdjustXY_2_1=here(db:utCurrentTool.tValue,world)
            db:jAdjustXY_2_1=herej()
            call db:updateTeachPos(db:pAdjustXY_2_1,db:bAdjustXY_2_1)
            call db:hmiAlert("First","info")
            call saveCall()
          endIf
          if db:utBtn_Bottom[2].Events.bClick==true
            db:utBtn_Bottom[2].Events.bClick=false
            //Press F3
            call moveRecPos("pAdjustXY_2_1")
          endIf
          if db:utBtn_Bottom[3].Events.bClick==true
            db:utBtn_Bottom[3].Events.bClick=false
            //Press F4
            switch db:utCurrentTool.nItem
              case 1
                if db:tTool2.trsf!={0,0,0,0,0,0}
                  call db:updateTool(2,false)
                else
                  call db:hmiAlert("CantSwitchTool2","warning")
                endIf
              break
              case 2
                call db:updateTool(1,false)
              break
            endSwitch
          endIf
          //
          if db:utBtn_Bottom[6].Events.bClick==true
            db:utBtn_Bottom[6].Events.bClick=false
            //Press F7
            resetMotion()
            db:utCtn_Message.Appearance.bVisibility=false
            db:nStep1=99
          endIf
          if db:utBtn_Bottom[7].Events.bClick==true
            db:utBtn_Bottom[7].Events.bClick=false
            //Press F8
            resetMotion()
            db:utCtn_Message.Appearance.bVisibility=false
            db:nStep1=20
          endIf
        break
        //
        case 20
          call db:updateStr(32,db:utLbl_Point.Common.sText,"Point：P2")
          call db:updateStr(42,db:utLbl_Step.Common.sText,"Step：2/2")
          //
          db:utImg_Example.Common.sSourceImage="images/6AxisAdjustXY2_2.png"

          //
          call db:updateTeachPos(db:pAdjustXY_2_2,db:bAdjustXY_2_2)
          //
          call db:updateBtn(85,"Reset,Here,Move,RZ+,RZ-,Calc.,Prev.,Done")
          //
          call db:updateInfo(101,db:utLbl_Info0.Data.nVal,db:utLbl_Info0.Common.sText,"0","Operation reminder：")
          call db:updateInfo(112,db:utLbl_Info1.Data.nVal,db:utLbl_Info1.Common.sText,"1","Press the RZ+(RZ-) & Move/Hold to rotate TCP 180°")
          call db:updateInfo(102,db:utLbl_Info2.Data.nVal,db:utLbl_Info2.Common.sText,"2","Touch to reference pointer in vertical attitude")
          call db:updateInfo(105,db:utLbl_Info3.Data.nVal,db:utLbl_Info3.Common.sText,"3","Press Here button to save the position")
          call db:updateInfo(104,db:utLbl_Info4.Data.nVal,db:utLbl_Info4.Common.sText,"4","Press Calc. button to get the TCP value")
          db:nStep1=21
        break
        //
        case 21
          if db:utBtn_Bottom[0].Events.bClick==true
            db:utBtn_Bottom[0].Events.bClick=false
            //Press F1
            call moveCalPos("GoBack_pAdjustXY_2_1")
          endIf
          if db:utBtn_Bottom[1].Events.bClick==true
            db:utBtn_Bottom[1].Events.bClick=false
            //Press F2
            db:bAdjustXY_2_2=true
            db:pAdjustXY_2_2=here(db:utCurrentTool.tValue,world)
            db:jAdjustXY_2_2=herej()
            call db:updateTeachPos(db:pAdjustXY_2_2,db:bAdjustXY_2_2)
            call db:hmiAlert("Second","info")
            call saveCall()
          endIf
          if db:utBtn_Bottom[2].Events.bClick==true
            db:utBtn_Bottom[2].Events.bClick=false
            //Press F3
            call moveRecPos("pAdjustXY_2_2")
          endIf
          if db:utBtn_Bottom[3].Events.bClick==true
            db:utBtn_Bottom[3].Events.bClick=false
            //Press F4
            call moveCalPos("Rz+180_pAdjustXY_2_1")
          endIf
          if db:utBtn_Bottom[4].Events.bClick==true
            db:utBtn_Bottom[4].Events.bClick=false
            //Press F5
            call moveCalPos("Rz-180_pAdjustXY_2_1")
          endIf
          if db:utBtn_Bottom[5].Events.bClick==true
            db:utBtn_Bottom[5].Events.bClick=false
            //Press F6
            call algorithm:CalAdjustXY2()
          endIf
          if db:utBtn_Bottom[6].Events.bClick==true
            db:utBtn_Bottom[6].Events.bClick=false
            //Press F7
            resetMotion()
            db:utCtn_Message.Appearance.bVisibility=false
            db:nStep1=10
          endIf
          if db:utBtn_Bottom[7].Events.bClick==true
            db:utBtn_Bottom[7].Events.bClick=false
            //Press F8
            resetMotion()
            db:utCtn_Message.Appearance.bVisibility=false
            db:nStep1=99
          endIf
        break
        //
        case 99
          db:utCtn_Function.Common.sSource="Page_Container_Main.html"
          //
          call db:updateBtn(83,"Null,Null,Null,Null,Null,Null,Null,Quit")
          //
          call db:updateInfo(99,db:utLbl_Info0.Data.nVal,db:utLbl_Info0.Common.sText,"0","")
          call db:updateInfo(99,db:utLbl_Info1.Data.nVal,db:utLbl_Info1.Common.sText,"1","")
          call db:updateInfo(100,db:utLbl_Info2.Data.nVal,db:utLbl_Info2.Common.sText,"0","TCP calibration application for TX2/TS2 robot")
          call db:updateInfo(99,db:utLbl_Info3.Data.nVal,db:utLbl_Info3.Common.sText,"3","")
          call db:updateInfo(99,db:utLbl_Info4.Data.nVal,db:utLbl_Info4.Common.sText,"4","")
          db:utBtn_Step[1].Events.bClick=false
          db:nStep1=10
        break
        //
      endSwitch
    endIf
    //**********************************************************************************************************************************
    //
    //**********************************************************************************************************************************
    //3点法修正TCP的XY
    if db:utImg_CheckBox_b[1].Data.bStatus==true
      switch db:nStep1
        case 10
          call db:updateStr(31,db:utLbl_Point.Common.sText,"Point：P1")
          call db:updateStr(43,db:utLbl_Step.Common.sText,"Step：1/3")
          //
          db:utImg_Example.Common.sSourceImage="images/6AxisAdjustXY3_1.png"

          //
          call db:updateTeachPos(db:pAdjustXY_3_1,db:bAdjustXY_3_1)
          //
          call db:updateBtn(84,"Align,Here,Move,Change,Null,Null,Prev.,Next")
          //
          call db:updateInfo(101,db:utLbl_Info0.Data.nVal,db:utLbl_Info0.Common.sText,"0","Operation reminder：")
          call db:updateInfo(114,db:utLbl_Info1.Data.nVal,db:utLbl_Info1.Common.sText,"1","Rotate TCP (RZ) close to middle position")
          call db:updateInfo(102,db:utLbl_Info2.Data.nVal,db:utLbl_Info2.Common.sText,"2","Touch to reference pointer in vertical attitude")
          call db:updateInfo(115,db:utLbl_Info3.Data.nVal,db:utLbl_Info3.Common.sText,"3","Ensure that the TCP(RZ) can be rotated ±60°")
          call db:updateInfo(105,db:utLbl_Info4.Data.nVal,db:utLbl_Info4.Common.sText,"4","Press Here button to save the position")
          //
          call db:updateTool(1,false)
          db:nStep1=11
        break
        //
        case 11
          if db:utBtn_Bottom[0].Events.bClick==true
            db:utBtn_Bottom[0].Events.bClick=false
            //Press F1
            call moveCalPos("Align")
          endIf
          if db:utBtn_Bottom[1].Events.bClick==true
            db:utBtn_Bottom[1].Events.bClick=false
            //Press F2
            db:bAdjustXY_3_1=true
            db:pAdjustXY_3_1=here(db:utCurrentTool.tValue,world)
            db:jAdjustXY_3_1=herej()
            call db:updateTeachPos(db:pAdjustXY_3_1,db:bAdjustXY_3_1)
            call db:hmiAlert("First","info")
            call saveCall()
          endIf
          if db:utBtn_Bottom[2].Events.bClick==true
            db:utBtn_Bottom[2].Events.bClick=false
            //Press F3
            call moveRecPos("pAdjustXY_3_1")
          endIf
          if db:utBtn_Bottom[3].Events.bClick==true
            db:utBtn_Bottom[3].Events.bClick=false
            //Press F4
            switch db:utCurrentTool.nItem
              case 1
                if db:tTool2.trsf!={0,0,0,0,0,0}
                  call db:updateTool(2,false)
                else
                  call db:hmiAlert("CantSwitchTool2","warning")
                endIf
              break
              case 2
                call db:updateTool(1,false)
              break
            endSwitch
          endIf
          if db:utBtn_Bottom[6].Events.bClick==true
            db:utBtn_Bottom[6].Events.bClick=false
            //Press F7
            resetMotion()
            db:utCtn_Message.Appearance.bVisibility=false
            db:nStep1=99
          endIf
          if db:utBtn_Bottom[7].Events.bClick==true
            db:utBtn_Bottom[7].Events.bClick=false
            //Press F8
            resetMotion()
            db:utCtn_Message.Appearance.bVisibility=false
            db:nStep1=20
          endIf
        break
        //
        case 20
          call db:updateStr(32,db:utLbl_Point.Common.sText,"Point：P2")
          call db:updateStr(44,db:utLbl_Step.Common.sText,"Step：2/3")
          //
          db:utImg_Example.Common.sSourceImage="images/6AxisAdjustXY3_2.png"

          //
          call db:updateTeachPos(db:pAdjustXY_3_2,db:bAdjustXY_3_2)
          //
          call db:updateBtn(86,"Reset,Here,Move,RZ+,Null,Null,Prev.,Next")
          //
          call db:updateInfo(101,db:utLbl_Info0.Data.nVal,db:utLbl_Info0.Common.sText,"0","Operation reminder：")
          call db:updateInfo(116,db:utLbl_Info1.Data.nVal,db:utLbl_Info1.Common.sText,"1","Press the RZ+ & Move/Hold to rotate TCP +60°")
          call db:updateInfo(102,db:utLbl_Info2.Data.nVal,db:utLbl_Info2.Common.sText,"2","Touch to reference pointer in vertical attitude")
          call db:updateInfo(105,db:utLbl_Info3.Data.nVal,db:utLbl_Info3.Common.sText,"3","Press Here button to save the position")
          call db:updateInfo(99,db:utLbl_Info4.Data.nVal,db:utLbl_Info4.Common.sText,"4","")
          //
          db:nStep1=21
        break
        //
        case 21
          if db:utBtn_Bottom[0].Events.bClick==true
            db:utBtn_Bottom[0].Events.bClick=false
            //Press F1
            call moveCalPos("GoBack_pAdjustXY_3_1")
          endIf
          if db:utBtn_Bottom[1].Events.bClick==true
            db:utBtn_Bottom[1].Events.bClick=false
            //Press F2
            db:bAdjustXY_3_2=true
            db:pAdjustXY_3_2=here(db:utCurrentTool.tValue,world)
            db:jAdjustXY_3_2=herej()
            call db:updateTeachPos(db:pAdjustXY_3_2,db:bAdjustXY_3_2)
            call db:hmiAlert("Second","info")
            call saveCall()
          endIf
          if db:utBtn_Bottom[2].Events.bClick==true
            db:utBtn_Bottom[2].Events.bClick=false
            //Press F3
            call moveRecPos("pAdjustXY_3_2")
          endIf
          if db:utBtn_Bottom[3].Events.bClick==true
            db:utBtn_Bottom[3].Events.bClick=false
            //Press F4
            call moveCalPos("Rz+60_pAdjustXY_3_1")
          endIf
          if db:utBtn_Bottom[6].Events.bClick==true
            db:utBtn_Bottom[6].Events.bClick=false
            //Press F7
            resetMotion()
            db:utCtn_Message.Appearance.bVisibility=false
            db:nStep1=10
          endIf
          if db:utBtn_Bottom[7].Events.bClick==true
            db:utBtn_Bottom[7].Events.bClick=false
            //Press F8
            resetMotion()
            db:utCtn_Message.Appearance.bVisibility=false
            db:nStep1=30
          endIf
        break
        //
        case 30
          call db:updateStr(33,db:utLbl_Point.Common.sText,"Point：P3")
          call db:updateStr(45,db:utLbl_Step.Common.sText,"Step：3/3")
          //
          db:utImg_Example.Common.sSourceImage="images/6AxisAdjustXY3_3.png"

          //
          call db:updateTeachPos(db:pAdjustXY_3_3,db:bAdjustXY_3_3)
          //
          call db:updateBtn(87,"Reset,Here,Move,RZ-,Null,Calc.,Prev.,Done")
          //
          call db:updateInfo(101,db:utLbl_Info0.Data.nVal,db:utLbl_Info0.Common.sText,"0","Operation reminder：")
          call db:updateInfo(117,db:utLbl_Info1.Data.nVal,db:utLbl_Info1.Common.sText,"1","Press the RZ+ & Move/Hold to rotate TCP -60°")
          call db:updateInfo(102,db:utLbl_Info2.Data.nVal,db:utLbl_Info2.Common.sText,"2","Touch to reference pointer in vertical attitude")
          call db:updateInfo(105,db:utLbl_Info3.Data.nVal,db:utLbl_Info3.Common.sText,"3","Press Here button to save the position")
          call db:updateInfo(104,db:utLbl_Info4.Data.nVal,db:utLbl_Info4.Common.sText,"4","Press Calc. button to get the TCP value")
          db:nStep1=31
        break
        //
        case 31
          if db:utBtn_Bottom[0].Events.bClick==true
            db:utBtn_Bottom[0].Events.bClick=false
            //Press F1
            call moveCalPos("GoBack_pAdjustXY_3_1")
          endIf
          if db:utBtn_Bottom[1].Events.bClick==true
            db:utBtn_Bottom[1].Events.bClick=false
            //Press F2
            db:bAdjustXY_3_3=true
            db:pAdjustXY_3_3=here(db:utCurrentTool.tValue,world)
            db:jAdjustXY_3_3=herej()
            call db:updateTeachPos(db:pAdjustXY_3_3,db:bAdjustXY_3_3)
            call db:hmiAlert("Third","info")
            call saveCall()
          endIf
          if db:utBtn_Bottom[2].Events.bClick==true
            db:utBtn_Bottom[2].Events.bClick=false
            //Press F3
            call moveRecPos("pAdjustXY_3_3")
          endIf
          if db:utBtn_Bottom[3].Events.bClick==true
            db:utBtn_Bottom[3].Events.bClick=false
            //Press F4
            call moveCalPos("Rz-60_pAdjustXY_3_1")
          endIf
          if db:utBtn_Bottom[5].Events.bClick==true
            db:utBtn_Bottom[5].Events.bClick=false
            //Press F6
            call algorithm:CalAdjustXY3()
          endIf
          if db:utBtn_Bottom[6].Events.bClick==true
            db:utBtn_Bottom[6].Events.bClick=false
            //Press F7
            resetMotion()
            db:utCtn_Message.Appearance.bVisibility=false
            db:nStep1=20
          endIf
          if db:utBtn_Bottom[7].Events.bClick==true
            db:utBtn_Bottom[7].Events.bClick=false
            //Press F8
            resetMotion()
            db:utCtn_Message.Appearance.bVisibility=false
            db:nStep1=99
          endIf
        break
        //
        case 99
          db:utCtn_Function.Common.sSource="Page_Container_Main.html"
          //
          call db:updateBtn(83,"Null,Null,Null,Null,Null,Null,Null,Quit")
          //
          call db:updateInfo(99,db:utLbl_Info0.Data.nVal,db:utLbl_Info0.Common.sText,"0","")
          call db:updateInfo(99,db:utLbl_Info1.Data.nVal,db:utLbl_Info1.Common.sText,"1","")
          call db:updateInfo(100,db:utLbl_Info2.Data.nVal,db:utLbl_Info2.Common.sText,"0","TCP calibration application for TX2/TS2 robot")
          call db:updateInfo(99,db:utLbl_Info3.Data.nVal,db:utLbl_Info3.Common.sText,"3","")
          call db:updateInfo(99,db:utLbl_Info4.Data.nVal,db:utLbl_Info4.Common.sText,"4","")
          db:utBtn_Step[1].Events.bClick=false
          db:nStep1=10
        break
        //
      endSwitch
    endIf
    //**********************************************************************************************************************************
  endIf
end

--- refreshBtn2_AdjZ.pgx ---
public program refreshBtn2_AdjZ()
begin
  if db:utBtn_Step[2].Events.bClick==true
    db:utCtn_Function.Common.sSource="Page_Container_Teach.html"
    //**********************************************************************************************************************************
    //2点法修正TCP的Z
    switch db:nStep2
      case 10
        call db:updateStr(31,db:utLbl_Point.Common.sText,"Point：P1")
        call db:updateStr(41,db:utLbl_Step.Common.sText,"Step：1/2")
        //
        db:utImg_Example.Common.sSourceImage="images/6AxisAdjustZ2_1.png"
        //
        call db:updateTeachPos(db:pAdjustZ_2_1,db:bAdjustZ_2_1)
        //
        call db:updateBtn(84,"Align,Here,Move,Change,Null,Null,Prev.,Next")
        //
        call db:updateInfo(101,db:utLbl_Info0.Data.nVal,db:utLbl_Info0.Common.sText,"0","Operation reminder：")
        call db:updateInfo(102,db:utLbl_Info1.Data.nVal,db:utLbl_Info1.Common.sText,"1","Touch to reference pointer in vertical attitude")
        call db:updateInfo(118,db:utLbl_Info2.Data.nVal,db:utLbl_Info2.Common.sText,"2","Ensure that the TCP(RX) or TCP(RY) can be rotated +60°")
        call db:updateInfo(105,db:utLbl_Info3.Data.nVal,db:utLbl_Info3.Common.sText,"3","Press Here button to save the position")
        call db:updateInfo(99,db:utLbl_Info4.Data.nVal,db:utLbl_Info4.Common.sText,"4","")
        //
        call db:updateTool(2,false)
        db:nStep2=11
      break
      //
      case 11
        if db:utBtn_Bottom[0].Events.bClick==true
          db:utBtn_Bottom[0].Events.bClick=false
          //Press F1
          call moveCalPos("Align")
        endIf
        if db:utBtn_Bottom[1].Events.bClick==true
          db:utBtn_Bottom[1].Events.bClick=false
          //Press F2
          db:bAdjustZ_2_1=true
          db:pAdjustZ_2_1=here(db:utCurrentTool.tValue,world)
          db:jAdjustZ_2_1=herej()
          call db:updateTeachPos(db:pAdjustZ_2_1,db:bAdjustZ_2_1)
          call db:hmiAlert("First","info")
          call saveCall()
        endIf
        if db:utBtn_Bottom[2].Events.bClick==true
          db:utBtn_Bottom[2].Events.bClick=false
          //Press F3
          call moveRecPos("pAdjustZ_2_1")
        endIf
        if db:utBtn_Bottom[3].Events.bClick==true
          db:utBtn_Bottom[3].Events.bClick=false
          //Press F4
          switch db:utCurrentTool.nItem
            case 2
              if db:tTool3.trsf!={0,0,0,0,0,0}
                call db:updateTool(3,false)
              else
                call db:hmiAlert("CantSwitchTool3","warning")
              endIf
            break
            case 3
              call db:updateTool(2,false)
            break
          endSwitch
        endIf
        //
        if db:utBtn_Bottom[6].Events.bClick==true
          db:utBtn_Bottom[6].Events.bClick=false
          //Press F7
          resetMotion()
          db:utCtn_Message.Appearance.bVisibility=false
          db:nStep2=99
        endIf
        if db:utBtn_Bottom[7].Events.bClick==true
          db:utBtn_Bottom[7].Events.bClick=false
          //Press F8
          resetMotion()
          db:utCtn_Message.Appearance.bVisibility=false
          db:nStep2=20
        endIf
      break
      //
      case 20
        call db:updateStr(32,db:utLbl_Point.Common.sText,"Point：P2")
        call db:updateStr(42,db:utLbl_Step.Common.sText,"Step：2/2")
        //
        db:utImg_Example.Common.sSourceImage="images/6AxisAdjustZ2_2.png"
        //
        call db:updateTeachPos(db:pAdjustZ_2_2,db:bAdjustZ_2_2)
        //
        call db:updateBtn(88,"Reset,Here,Move,RX+,RY+,Calc.,Prev.,Done")
        //
        call db:updateInfo(101,db:utLbl_Info0.Data.nVal,db:utLbl_Info0.Common.sText,"0","Operation reminder：")
        call db:updateInfo(119,db:utLbl_Info1.Data.nVal,db:utLbl_Info1.Common.sText,"1","Press the RX+(RY+) & Move/Hold to rotate TCP 60°")
        call db:updateInfo(120,db:utLbl_Info2.Data.nVal,db:utLbl_Info2.Common.sText,"2","Touch to reference pointer in current attitude")
        call db:updateInfo(105,db:utLbl_Info3.Data.nVal,db:utLbl_Info3.Common.sText,"3","Press Here button to save the position")
        call db:updateInfo(104,db:utLbl_Info4.Data.nVal,db:utLbl_Info4.Common.sText,"4","Press Calc. button to get the TCP value")
        db:nStep2=21
      break
      //
      case 21
        if db:utBtn_Bottom[0].Events.bClick==true
          db:utBtn_Bottom[0].Events.bClick=false
          //Press F1
          call moveCalPos("GoBack_pAdjustZ_2_1")
        endIf
        if db:utBtn_Bottom[1].Events.bClick==true
          db:utBtn_Bottom[1].Events.bClick=false
          //Press F2
          db:bAdjustZ_2_2=true
          db:pAdjustZ_2_2=here(db:utCurrentTool.tValue,world)
          db:jAdjustZ_2_2=herej()
          call db:updateTeachPos(db:pAdjustZ_2_2,db:bAdjustZ_2_2)
          call db:hmiAlert("Second","info")
          call saveCall()
        endIf
        if db:utBtn_Bottom[2].Events.bClick==true
          db:utBtn_Bottom[2].Events.bClick=false
          //Press F3
          call moveRecPos("pAdjustZ_2_2")
        endIf
        if db:utBtn_Bottom[3].Events.bClick==true
          db:utBtn_Bottom[3].Events.bClick=false
          //Press F4
          call moveCalPos("Rx+60_pAdjustZ_2_1")
        endIf
        if db:utBtn_Bottom[4].Events.bClick==true
          db:utBtn_Bottom[4].Events.bClick=false
          //Press F5
          call moveCalPos("Ry+60_pAdjustZ_2_1")
        endIf
        if db:utBtn_Bottom[5].Events.bClick==true
          db:utBtn_Bottom[5].Events.bClick=false
          //Press F6
          call algorithm:CalAdjustZ()
        endIf
        if db:utBtn_Bottom[6].Events.bClick==true
          db:utBtn_Bottom[6].Events.bClick=false
          //Press F7
          resetMotion()
          db:utCtn_Message.Appearance.bVisibility=false
          db:nStep2=10
        endIf
        if db:utBtn_Bottom[7].Events.bClick==true
          db:utBtn_Bottom[7].Events.bClick=false
          //Press F8
          resetMotion()
          db:utCtn_Message.Appearance.bVisibility=false
          db:nStep2=99
        endIf
      break
      //
      case 99
        db:utCtn_Function.Common.sSource="Page_Container_Main.html"
        //
        call db:updateBtn(83,"Null,Null,Null,Null,Null,Null,Null,Quit")
        //
        call db:updateInfo(99,db:utLbl_Info0.Data.nVal,db:utLbl_Info0.Common.sText,"0","")
        call db:updateInfo(99,db:utLbl_Info1.Data.nVal,db:utLbl_Info1.Common.sText,"1","")
        call db:updateInfo(100,db:utLbl_Info2.Data.nVal,db:utLbl_Info2.Common.sText,"0","TCP calibration application for TX2/TS2 robot")
        call db:updateInfo(99,db:utLbl_Info3.Data.nVal,db:utLbl_Info3.Common.sText,"3","")
        call db:updateInfo(99,db:utLbl_Info4.Data.nVal,db:utLbl_Info4.Common.sText,"4","")
        db:utBtn_Step[2].Events.bClick=false
        db:nStep2=10
      break
      //
    endSwitch
    //**********************************************************************************************************************************
  endIf
end

--- refreshBtn3_Test.pgx ---
public program refreshBtn3_Test()
  local num l_nStep
  local bool l_bOut
  local bool l_bTaskStatusErr
  local num l_nI
begin
  if db:utBtn_Step[3].Events.bClick==true
    db:utCtn_Function.Common.sSource="Page_Container_Test.html"
    //**********************************************************************************************************************************
    switch db:nStep3
      case 10
        call db:updateBtn(89,"Align,Here,Move,Change,Null,Null,Prev.,Next")
        //
        call db:updateTool(db:utCurrentTool.nItem,true)
        //
        db:utLbl_ToolValue_Data[0].Common.sText=toString(".3",db:utCurrentTool.tValue.trsf.x)
        db:utLbl_ToolValue_Data[1].Common.sText=toString(".3",db:utCurrentTool.tValue.trsf.y)
        db:utLbl_ToolValue_Data[2].Common.sText=toString(".3",db:utCurrentTool.tValue.trsf.z)
        db:utLbl_ToolValue_Data[3].Common.sText=toString(".3",db:utCurrentTool.tValue.trsf.rx)
        db:utLbl_ToolValue_Data[4].Common.sText=toString(".3",db:utCurrentTool.tValue.trsf.ry)
        db:utLbl_ToolValue_Data[5].Common.sText=toString(".3",db:utCurrentTool.tValue.trsf.rz)
        //
        db:utTxt_OffsetValue_Data[0].Common.nValue=round(db:trOffset.x*1000)/1000
        db:utTxt_OffsetValue_Data[1].Common.nValue=round(db:trOffset.y*1000)/1000
        db:utTxt_OffsetValue_Data[2].Common.nValue=round(db:trOffset.z*1000)/1000
        db:utTxt_OffsetValue_Data[3].Common.nValue=round(db:trOffset.rx*1000)/1000
        db:utTxt_OffsetValue_Data[4].Common.nValue=round(db:trOffset.ry*1000)/1000
        db:utTxt_OffsetValue_Data[5].Common.nValue=round(db:trOffset.rz*1000)/1000
        db:nStep3=20
      break
      //
      case 20
        //**********************************************************************************************************************************
        //刷新当前工具值
        if db:utCurrentTool.nItem!=db:utCurrentTool.nItemM or db:bRefresh==true
          db:utCurrentTool.nItemM=db:utCurrentTool.nItem
          db:bRefresh=false
          call db:updateTool(db:utCurrentTool.nItem,true)
        db:utLbl_ToolValue_Data[0].Common.sText=toString(".3",db:utCurrentTool.tValue.trsf.x)
        db:utLbl_ToolValue_Data[1].Common.sText=toString(".3",db:utCurrentTool.tValue.trsf.y)
        db:utLbl_ToolValue_Data[2].Common.sText=toString(".3",db:utCurrentTool.tValue.trsf.z)
        db:utLbl_ToolValue_Data[3].Common.sText=toString(".3",db:utCurrentTool.tValue.trsf.rx)
        db:utLbl_ToolValue_Data[4].Common.sText=toString(".3",db:utCurrentTool.tValue.trsf.ry)
        db:utLbl_ToolValue_Data[5].Common.sText=toString(".3",db:utCurrentTool.tValue.trsf.rz)
        endIf
        //刷新当前工具序号（Previous）
        if db:utImg_Previous.Events.bClick==true
          db:utImg_Previous.Events.bClick=false
          switch db:utCurrentTool.nItem
            case 1,2,3
              db:utCurrentTool.nItem=db:utCurrentTool.nItem-1
            break
            case 0
              db:utCurrentTool.nItem=3
            break
            default
              db:utCurrentTool.nItem=0
            break
          endSwitch
        endIf
        //刷新当前工具序号（Next）
        if db:utImg_Next.Events.bClick==true
          db:utImg_Next.Events.bClick=false
          switch db:utCurrentTool.nItem
            case 0,1,2
              db:utCurrentTool.nItem=db:utCurrentTool.nItem+1
            break
            case 3
              db:utCurrentTool.nItem=0
            break
            default
              db:utCurrentTool.nItem=0
            break
          endSwitch
        endIf

        //**********************************************************************************************************************************
        //
        //
        //**********************************************************************************************************************************
        //刷新当前偏移值
        l_nStep=0
        l_bOut=false
        do
          switch l_nStep
            case 0
              if db:utTxt_OffsetValue_Data[0].Common.nValue==db:trOffset.x
                l_nStep=1
              else
                l_nStep=99
              endIf
            break
            case 1
              if db:utTxt_OffsetValue_Data[1].Common.nValue==db:trOffset.y
                l_nStep=2
              else
                l_nStep=99
              endIf
            break
            case 2
              if db:utTxt_OffsetValue_Data[2].Common.nValue==db:trOffset.z
                l_nStep=3
              else
                l_nStep=99
              endIf
            break
            case 3
              if db:utTxt_OffsetValue_Data[3].Common.nValue==db:trOffset.rx
                l_nStep=4
              else
                l_nStep=99
              endIf
            break
            case 4
              if db:utTxt_OffsetValue_Data[4].Common.nValue==db:trOffset.ry
                l_nStep=5
              else
                l_nStep=99
              endIf
            break
            case 5
              if db:utTxt_OffsetValue_Data[5].Common.nValue==db:trOffset.rz
                l_nStep=100
              else
                l_nStep=99
              endIf
            break
            case 99
              db:utTxt_OffsetValue_Data[0].Common.nValue=round(db:utTxt_OffsetValue_Data[0].Common.nValue*1000)/1000
              db:utTxt_OffsetValue_Data[1].Common.nValue=round(db:utTxt_OffsetValue_Data[1].Common.nValue*1000)/1000
              db:utTxt_OffsetValue_Data[2].Common.nValue=round(db:utTxt_OffsetValue_Data[2].Common.nValue*1000)/1000
              db:utTxt_OffsetValue_Data[3].Common.nValue=round(db:utTxt_OffsetValue_Data[3].Common.nValue*1000)/1000
              db:utTxt_OffsetValue_Data[4].Common.nValue=round(db:utTxt_OffsetValue_Data[4].Common.nValue*1000)/1000
              db:utTxt_OffsetValue_Data[5].Common.nValue=round(db:utTxt_OffsetValue_Data[5].Common.nValue*1000)/1000
              //
              db:trOffset.x=db:utTxt_OffsetValue_Data[0].Common.nValue
              db:trOffset.y=db:utTxt_OffsetValue_Data[1].Common.nValue
              db:trOffset.z=db:utTxt_OffsetValue_Data[2].Common.nValue
              db:trOffset.rx=db:utTxt_OffsetValue_Data[3].Common.nValue
              db:trOffset.ry=db:utTxt_OffsetValue_Data[4].Common.nValue
              db:trOffset.rz=db:utTxt_OffsetValue_Data[5].Common.nValue
              //
              db:bRefresh=true
              l_bOut=true
            break
            case 100
              l_bOut=true
            break
          endSwitch
        until l_bOut
        //**********************************************************************************************************************************
        if db:utImg_Switch.Events.bClick==true
          db:utImg_Switch.Events.bClick=false
          if db:utImg_Switch.Data.bStatus==false
            db:utImg_Switch.Common.sSourceImage=db:utImg_Switch.Data.sSourceImg1
            db:utImg_Switch.Data.bStatus=true
            db:bRefresh=true
            for l_nI=0 to 5
              db:utTxt_OffsetValue_Data[l_nI].Appearance.sBackgroundColour="#7CFA3F"
            endFor
          else
            db:utImg_Switch.Common.sSourceImage=db:utImg_Switch.Data.sSourceImg2
            db:utImg_Switch.Data.bStatus=false
            db:bRefresh=true
            for l_nI=0 to 5
              db:utTxt_OffsetValue_Data[l_nI].Appearance.sBackgroundColour="#EEFF00"
            endFor
          endIf
        endIf
        //**********************************************************************************************************************************
        if db:utBtn_Bottom[0].Events.bClick==true
          db:utBtn_Bottom[0].Events.bClick=false
          //Press F1
          call moveCalPos("Align")
        endIf
        //
        if db:utBtn_Bottom[7].Events.bClick==true
          db:utBtn_Bottom[7].Events.bClick=false
          //Press F8
          db:utCtn_Function.Common.sSource="Page_Container_Main.html"
          //
          call db:updateBtn(83,"Null,Null,Null,Null,Null,Null,Null,Quit")
          //
          call db:updateInfo(99,db:utLbl_Info0.Data.nVal,db:utLbl_Info0.Common.sText,"0","")
          call db:updateInfo(99,db:utLbl_Info1.Data.nVal,db:utLbl_Info1.Common.sText,"1","")
          call db:updateInfo(100,db:utLbl_Info2.Data.nVal,db:utLbl_Info2.Common.sText,"0","TCP calibration application for TX2/TS2 robot")
          call db:updateInfo(99,db:utLbl_Info3.Data.nVal,db:utLbl_Info3.Common.sText,"3","")
          call db:updateInfo(99,db:utLbl_Info4.Data.nVal,db:utLbl_Info4.Common.sText,"4","")
          db:utBtn_Step[3].Events.bClick=false
          db:nStep3=10
          resetMotion()
          db:utCtn_Message.Appearance.bVisibility=false
        endIf
      break
    endSwitch
  endIf

end

--- saveCall.pgx ---
program saveCall()
begin
  if taskStatus("Save")==-1
    taskCreate "Save",100,saveTask()
  endIf
end

--- saveTask.pgx ---
program saveTask()
begin
  db:libSave()
end

--- stop.pgx ---
program stop()
begin



end
